Fanuc KAREL source: KO00118.KL

PROGRAM KO00118
%NOLOCKGROUP
VAR
  A: ARRAY[2] OF BYTE
  B: ARRAY[2] OF BYTE
  OUT: REAL
BEGIN
  A[1] = 1
  B[1] = 2
  OUT = ATAN2(A[1], B[1])
END KO00118
